// Én rute i kartet. x teller østover og y nordover fra kartets origo, som i verden.
TYPE GridCell :
STRUCT
	x : DINT;
	y : DINT;
END_STRUCT
END_TYPE

(* stored: Version 1.1.0.1, ProductVersion 3.1.4026.12
   DUT GridCell: Id {0a0df2dd-0c72-4488-b025-27794f2f03af} *)
